Fanuc KAREL source: ka00131.KL

-- PROVISIONAL review KL for V770-1; original PC SHA256 5313788d550a2d6cc4ce234ad17aa5d5bf2dcfb67c1255c89085ff3eab12156a
-- Incomplete behavior may be omitted. Consult companion uncertainty JSON. Do not deploy.
PROGRAM KA00131
%NOLOCKGROUP
-- UNRESOLVED_DECL SRC type=002018
-- UNRESOLVED_DECL DST type=002018
BEGIN
  -- UNRESOLVED_PC offsets 5-19; opcodes 2E,22,9D,33,B2
  -- UNRESOLVED_PC offsets 24-42; opcodes 22,9D,33,B1,22,9D,33,B2
  -- UNRESOLVED_PC offsets 47-51; opcodes 7F
END KA00131
